(* IEC 61131-3 sources: SRCI_CLIENT_PLC/RobotLibrary/Library/Structures/Dynamics, 3 files *)

(* ---- DefaultDynamics.st ---- *)
{attribute 'pack_mode' := '1'}
// -------------------------------------------------------------------------
//  SRCI Robot Library
// -------------------------------------------------------------------------
//
//  Object:      DefaultDynamics
//  Author:      Thorsten Brach
//  Date:        2024-06-01
//
//  Description:
//
//
//  Copyright:
//    (C) 2024 Thorsten Brach. All rights reserved
//             Licensed under the MIT License.
//
//  Disclaimer:
//    This project is provided without any guarantee and can be used for
//    private and commercial purposes. Any use is at the user’s
//    own risk and responsibility.
//
// -------------------------------------------------------------------------
TYPE DefaultDynamics :
STRUCT
  /// Timestamp
  Timestamp        : IEC_TIMESTAMP;
  /// Maximum velocity for the axes.
  /// Range [%]:
  /// •  <0% : Use default velocity given by the user
  /// •   0% : Use internal minimal velocity
  /// • 100% : Use the entire reference velocity, given by the user
  VelocityRate     : REAL;
  /// Maximum acceleration.
  /// Range [%]:
  /// •  <0% : Use default acceleration given by the user
  /// •   0% : Use internal minimal acceleration
  /// • 100% : Use the entire reference acceleration, given by the user
  AccelerationRate : REAL;
  /// Maximum deceleration.
  /// Range [%] :
  /// •  <0% : Use default deceleration given by the user
  /// •   0% : Use internal minimal deceleration
  /// • 100% : Use the entire reference deceleration, given by the user
  DecelerationRate : REAL;
  /// Maximum jerk
  /// Range [%] :
  /// •  <0% : Use default jerk given by the user
  /// •   0% : Use internal minimal jerk
  /// • 100% : Use the entire reference jerk, given by the user (Trapezoidal if possible)
  JerkRate         : REAL;
END_STRUCT
END_TYPE

(* ---- ReferenceDynamics.st ---- *)
{attribute 'pack_mode' := '1'}
// -------------------------------------------------------------------------
//  SRCI Robot Library
// -------------------------------------------------------------------------
//
//  Object:      ReferenceDynamics
//  Author:      Thorsten Brach
//  Date:        2024-06-01
//
//  Description:
//
//
//  Copyright:
//    (C) 2024 Thorsten Brach. All rights reserved
//             Licensed under the MIT License.
//
//  Disclaimer:
//    This project is provided without any guarantee and can be used for
//    private and commercial purposes. Any use is at the user’s
//    own risk and responsibility.
//
// -------------------------------------------------------------------------
TYPE ReferenceDynamics :
STRUCT
  /// Timestamp
  Timestamp             : IEC_TIMESTAMP;
  /// Path velocity [mm/s](tangent) at 100%
  /// • <0: (default) - Do not change values
  /// • ≥0: Change values according to input value
  VelocityReference     : REAL;
  /// Path acceleration [mm/s2] at 100%
  /// • <0: (default) - Do not change values
  /// • ≥0: Change values according to input value
  AccelerationReference : REAL;
  /// Path deceleration [mm/s2] at 100%
  /// • <0: (default) - Do not change values
  /// • ≥0: Change values according to input value
  DecelerationReference : REAL;
  /// Jerk [mm/s3] at 100%
  /// • <0: (default) - Do not change values
  /// • ≥0: Change values according to input value
  JerkReference        : REAL;
END_STRUCT
END_TYPE

(* ---- RobotDynamics.st ---- *)
{attribute 'pack_mode' := '1'}
// -------------------------------------------------------------------------
//  SRCI Robot Library
// -------------------------------------------------------------------------
//
//  Object:      RobotDynamics
//  Author:      Thorsten Brach
//  Date:        2025-10-15
//
//  Description:
//
//
//  Copyright:
//    (C) 2025 Thorsten Brach. All rights reserved
//             Licensed under the MIT License.
//
//  Disclaimer:
//    This project is provided without any guarantee and can be used for
//    private and commercial purposes. Any use is at the user’s
//    own risk and responsibility.
//
// -------------------------------------------------------------------------
TYPE RobotDynamics :
STRUCT
  /// TCP velocity in % of nominal velocity
  /// •  <0% (default) o Use default velocity
  /// •   0%           o Use internal minimal velocity
  /// • 100%           o Use maximal reference velocity
  /// See chapter 5.5.7 Robot dynamics
  VelocityRate     : REAL;
  /// Acceleration for movement in % of nominal acceleration
  /// •  <0% (default) o Use default acceleration
  /// •   0%           o Use internal minimal acceleration
  /// • 100%:          o Use maximal reference acceleration
  /// See chapter 5.5.7 Robot dynamics
  AccelerationRate : REAL;
  /// Deceleration for movement in % of nominal deceleration
  /// •  <0% (default) o Use default deceleration
  /// •   0%           o Use internal minimal deceleration
  /// • 100%           o Use maximal reference deceleration
  /// See chapter 5.5.7 Robot dynamics
  DecelerationRate : REAL;
  /// Jerk of the movement in % of nominal jerk
  /// •  <0% (default) o Use default jerk
  /// •   0%           o Use internal minimal jerk
  /// • 100%           o Use maximal reference jerk
  /// See chapter 5.5.7 Robot dynamics
  JerkRate         : REAL;
END_STRUCT
END_TYPE
